(* IEC 61131-3 sources: STAR-PLC-Agent/results/raw/four_group_20261114/star_deepseek_v4/SELF004/generation/sim_00, 1 file *)

(* ---- test_program.st ---- *)
PROGRAM PLC_PRG
VAR
 BenchStep : UDINT := 0;
 BenchCalls : UDINT := 0;
 BenchDone : BOOL := FALSE;
 BenchUut0 : FB_Task;
 BenchUut1 : FB_Task;
 TraceIn_Start : ARRAY[0..13] OF BOOL;
 TraceIn_Stop : ARRAY[0..13] OF BOOL;
 TraceIn_AtExit : ARRAY[0..13] OF BOOL;
 TraceIn_Jam : ARRAY[0..13] OF BOOL;
 TraceIn_Reset : ARRAY[0..13] OF BOOL;
 TraceOut_Belt : ARRAY[0..13] OF BOOL;
 TraceOut_Complete : ARRAY[0..13] OF BOOL;
 TraceOut_Fault : ARRAY[0..13] OF BOOL;
END_VAR

IF NOT BenchDone THEN
 CASE BenchStep OF
 0:
   BenchUut0.Start := TRUE;
   BenchUut0.Stop := FALSE;
   BenchUut0.AtExit := TRUE;
   BenchUut0.Jam := FALSE;
   BenchUut0.Reset := FALSE;
   TraceIn_Start[0] := BenchUut0.Start;
   TraceIn_Stop[0] := BenchUut0.Stop;
   TraceIn_AtExit[0] := BenchUut0.AtExit;
   TraceIn_Jam[0] := BenchUut0.Jam;
   TraceIn_Reset[0] := BenchUut0.Reset;
   BenchUut0();
   TraceOut_Belt[0] := BenchUut0.Belt;
   TraceOut_Complete[0] := BenchUut0.Complete;
   TraceOut_Fault[0] := BenchUut0.Fault;
   BenchCalls := BenchCalls + 1;
 1:
   BenchUut0.Start := TRUE;
   BenchUut0.Stop := FALSE;
   BenchUut0.AtExit := FALSE;
   BenchUut0.Jam := FALSE;
   BenchUut0.Reset := FALSE;
   TraceIn_Start[1] := BenchUut0.Start;
   TraceIn_Stop[1] := BenchUut0.Stop;
   TraceIn_AtExit[1] := BenchUut0.AtExit;
   TraceIn_Jam[1] := BenchUut0.Jam;
   TraceIn_Reset[1] := BenchUut0.Reset;
   BenchUut0();
   TraceOut_Belt[1] := BenchUut0.Belt;
   TraceOut_Complete[1] := BenchUut0.Complete;
   TraceOut_Fault[1] := BenchUut0.Fault;
   BenchCalls := BenchCalls + 1;
 2:
   BenchUut0.Start := FALSE;
   BenchUut0.Stop := FALSE;
   BenchUut0.AtExit := FALSE;
   BenchUut0.Jam := FALSE;
   BenchUut0.Reset := FALSE;
   TraceIn_Start[2] := BenchUut0.Start;
   TraceIn_Stop[2] := BenchUut0.Stop;
   TraceIn_AtExit[2] := BenchUut0.AtExit;
   TraceIn_Jam[2] := BenchUut0.Jam;
   TraceIn_Reset[2] := BenchUut0.Reset;
   BenchUut0();
   TraceOut_Belt[2] := BenchUut0.Belt;
   TraceOut_Complete[2] := BenchUut0.Complete;
   TraceOut_Fault[2] := BenchUut0.Fault;
   BenchCalls := BenchCalls + 1;
 3:
   BenchUut0.Start := FALSE;
   BenchUut0.Stop := FALSE;
   BenchUut0.AtExit := TRUE;
   BenchUut0.Jam := FALSE;
   BenchUut0.Reset := FALSE;
   TraceIn_Start[3] := BenchUut0.Start;
   TraceIn_Stop[3] := BenchUut0.Stop;
   TraceIn_AtExit[3] := BenchUut0.AtExit;
   TraceIn_Jam[3] := BenchUut0.Jam;
   TraceIn_Reset[3] := BenchUut0.Reset;
   BenchUut0();
   TraceOut_Belt[3] := BenchUut0.Belt;
   TraceOut_Complete[3] := BenchUut0.Complete;
   TraceOut_Fault[3] := BenchUut0.Fault;
   BenchCalls := BenchCalls + 1;
 4:
   BenchUut0.Start := TRUE;
   BenchUut0.Stop := FALSE;
   BenchUut0.AtExit := FALSE;
   BenchUut0.Jam := FALSE;
   BenchUut0.Reset := FALSE;
   TraceIn_Start[4] := BenchUut0.Start;
   TraceIn_Stop[4] := BenchUut0.Stop;
   TraceIn_AtExit[4] := BenchUut0.AtExit;
   TraceIn_Jam[4] := BenchUut0.Jam;
   TraceIn_Reset[4] := BenchUut0.Reset;
   BenchUut0();
   TraceOut_Belt[4] := BenchUut0.Belt;
   TraceOut_Complete[4] := BenchUut0.Complete;
   TraceOut_Fault[4] := BenchUut0.Fault;
   BenchCalls := BenchCalls + 1;
 5:
   BenchUut0.Start := FALSE;
   BenchUut0.Stop := TRUE;
   BenchUut0.AtExit := FALSE;
   BenchUut0.Jam := FALSE;
   BenchUut0.Reset := FALSE;
   TraceIn_Start[5] := BenchUut0.Start;
   TraceIn_Stop[5] := BenchUut0.Stop;
   TraceIn_AtExit[5] := BenchUut0.AtExit;
   TraceIn_Jam[5] := BenchUut0.Jam;
   TraceIn_Reset[5] := BenchUut0.Reset;
   BenchUut0();
   TraceOut_Belt[5] := BenchUut0.Belt;
   TraceOut_Complete[5] := BenchUut0.Complete;
   TraceOut_Fault[5] := BenchUut0.Fault;
   BenchCalls := BenchCalls + 1;
 6:
   BenchUut0.Start := FALSE;
   BenchUut0.Stop := FALSE;
   BenchUut0.AtExit := FALSE;
   BenchUut0.Jam := FALSE;
   BenchUut0.Reset := FALSE;
   TraceIn_Start[6] := BenchUut0.Start;
   TraceIn_Stop[6] := BenchUut0.Stop;
   TraceIn_AtExit[6] := BenchUut0.AtExit;
   TraceIn_Jam[6] := BenchUut0.Jam;
   TraceIn_Reset[6] := BenchUut0.Reset;
   BenchUut0();
   TraceOut_Belt[6] := BenchUut0.Belt;
   TraceOut_Complete[6] := BenchUut0.Complete;
   TraceOut_Fault[6] := BenchUut0.Fault;
   BenchCalls := BenchCalls + 1;
 7:
   BenchUut1.Start := TRUE;
   BenchUut1.Stop := FALSE;
   BenchUut1.AtExit := FALSE;
   BenchUut1.Jam := TRUE;
   BenchUut1.Reset := TRUE;
   TraceIn_Start[7] := BenchUut1.Start;
   TraceIn_Stop[7] := BenchUut1.Stop;
   TraceIn_AtExit[7] := BenchUut1.AtExit;
   TraceIn_Jam[7] := BenchUut1.Jam;
   TraceIn_Reset[7] := BenchUut1.Reset;
   BenchUut1();
   TraceOut_Belt[7] := BenchUut1.Belt;
   TraceOut_Complete[7] := BenchUut1.Complete;
   TraceOut_Fault[7] := BenchUut1.Fault;
   BenchCalls := BenchCalls + 1;
 8:
   BenchUut1.Start := FALSE;
   BenchUut1.Stop := FALSE;
   BenchUut1.AtExit := FALSE;
   BenchUut1.Jam := FALSE;
   BenchUut1.Reset := FALSE;
   TraceIn_Start[8] := BenchUut1.Start;
   TraceIn_Stop[8] := BenchUut1.Stop;
   TraceIn_AtExit[8] := BenchUut1.AtExit;
   TraceIn_Jam[8] := BenchUut1.Jam;
   TraceIn_Reset[8] := BenchUut1.Reset;
   BenchUut1();
   TraceOut_Belt[8] := BenchUut1.Belt;
   TraceOut_Complete[8] := BenchUut1.Complete;
   TraceOut_Fault[8] := BenchUut1.Fault;
   BenchCalls := BenchCalls + 1;
 9:
   BenchUut1.Start := FALSE;
   BenchUut1.Stop := FALSE;
   BenchUut1.AtExit := FALSE;
   BenchUut1.Jam := FALSE;
   BenchUut1.Reset := TRUE;
   TraceIn_Start[9] := BenchUut1.Start;
   TraceIn_Stop[9] := BenchUut1.Stop;
   TraceIn_AtExit[9] := BenchUut1.AtExit;
   TraceIn_Jam[9] := BenchUut1.Jam;
   TraceIn_Reset[9] := BenchUut1.Reset;
   BenchUut1();
   TraceOut_Belt[9] := BenchUut1.Belt;
   TraceOut_Complete[9] := BenchUut1.Complete;
   TraceOut_Fault[9] := BenchUut1.Fault;
   BenchCalls := BenchCalls + 1;
 10:
   BenchUut1.Start := TRUE;
   BenchUut1.Stop := FALSE;
   BenchUut1.AtExit := FALSE;
   BenchUut1.Jam := FALSE;
   BenchUut1.Reset := FALSE;
   TraceIn_Start[10] := BenchUut1.Start;
   TraceIn_Stop[10] := BenchUut1.Stop;
   TraceIn_AtExit[10] := BenchUut1.AtExit;
   TraceIn_Jam[10] := BenchUut1.Jam;
   TraceIn_Reset[10] := BenchUut1.Reset;
   BenchUut1();
   TraceOut_Belt[10] := BenchUut1.Belt;
   TraceOut_Complete[10] := BenchUut1.Complete;
   TraceOut_Fault[10] := BenchUut1.Fault;
   BenchCalls := BenchCalls + 1;
 11:
   BenchUut1.Start := FALSE;
   BenchUut1.Stop := FALSE;
   BenchUut1.AtExit := FALSE;
   BenchUut1.Jam := TRUE;
   BenchUut1.Reset := FALSE;
   TraceIn_Start[11] := BenchUut1.Start;
   TraceIn_Stop[11] := BenchUut1.Stop;
   TraceIn_AtExit[11] := BenchUut1.AtExit;
   TraceIn_Jam[11] := BenchUut1.Jam;
   TraceIn_Reset[11] := BenchUut1.Reset;
   BenchUut1();
   TraceOut_Belt[11] := BenchUut1.Belt;
   TraceOut_Complete[11] := BenchUut1.Complete;
   TraceOut_Fault[11] := BenchUut1.Fault;
   BenchCalls := BenchCalls + 1;
 12:
   BenchUut1.Start := TRUE;
   BenchUut1.Stop := FALSE;
   BenchUut1.AtExit := FALSE;
   BenchUut1.Jam := TRUE;
   BenchUut1.Reset := TRUE;
   TraceIn_Start[12] := BenchUut1.Start;
   TraceIn_Stop[12] := BenchUut1.Stop;
   TraceIn_AtExit[12] := BenchUut1.AtExit;
   TraceIn_Jam[12] := BenchUut1.Jam;
   TraceIn_Reset[12] := BenchUut1.Reset;
   BenchUut1();
   TraceOut_Belt[12] := BenchUut1.Belt;
   TraceOut_Complete[12] := BenchUut1.Complete;
   TraceOut_Fault[12] := BenchUut1.Fault;
   BenchCalls := BenchCalls + 1;
 13:
   BenchUut1.Start := FALSE;
   BenchUut1.Stop := FALSE;
   BenchUut1.AtExit := FALSE;
   BenchUut1.Jam := FALSE;
   BenchUut1.Reset := TRUE;
   TraceIn_Start[13] := BenchUut1.Start;
   TraceIn_Stop[13] := BenchUut1.Stop;
   TraceIn_AtExit[13] := BenchUut1.AtExit;
   TraceIn_Jam[13] := BenchUut1.Jam;
   TraceIn_Reset[13] := BenchUut1.Reset;
   BenchUut1();
   TraceOut_Belt[13] := BenchUut1.Belt;
   TraceOut_Complete[13] := BenchUut1.Complete;
   TraceOut_Fault[13] := BenchUut1.Fault;
   BenchCalls := BenchCalls + 1;
 END_CASE;
 BenchStep := BenchStep + 1;
 IF BenchStep >= 14 THEN BenchDone := TRUE; END_IF;
END_IF;
END_PROGRAM
